Fanuc KAREL source: KT00230.KL

PROGRAM KT00230
%NOLOCKGROUP
VAR
  B1: BOOLEAN
  Y2: ARRAY[2] OF BYTE
  OUT: INTEGER
BEGIN
  B1 = TRUE
    Y2[1] = 3
  OUT = B1 OR Y2[1]
END KT00230
